// RUN: sclang-gen --emit=ast %s | FileCheck %s

function f : int
var_temp
  x : int;
end_var
begin
  x := 3;
  case x of
    1..3: x := 10;
    5, 7..8: x := 20;
  else
    x := 30;
  end_case;
end_function

// CHECK: CaseLabel
// CHECK: CaseLabel
